// HMI -> PLC: commands of the screen Main.
TYPE ST_HMI_SystemCommand :
STRUCT
    bResetAll : BOOL;  // Tap - reset of all devices of this system (evaluated on the rising edge)
END_STRUCT
END_TYPE

(* stored: Version 1.1.0.1
   DUT ST_HMI_SystemCommand: Id {faa143dc-fd00-4930-8e2a-f7ec609b33dd} *)
